(* IEC 61131-3 sources: PLC-Static-Analysis/modules/plc-rules/src/test/resources/PLCA-L008, 2 files *)

(* ---- compliant.st ---- *)
PROGRAM P_L008ok
VAR
    n : INT;
    m : INT;
    r : REAL;
    b : BOOL;
    c : BOOL;
    q : BOOL;
END_VAR
IF n > 10 THEN
    n := n - 20;
    IF n > 5 THEN
        q := TRUE;
    END_IF
END_IF
FOR m := 1 TO 10 DO
    IF n > 10 THEN
        q := TRUE;
    END_IF
    n := n + 1;
END_FOR
IF n > 10 THEN
    IF n > 50 THEN
        q := TRUE;
    END_IF
END_IF
END_PROGRAM

(* ---- noncompliant.st ---- *)
PROGRAM P_L008
VAR
    n : INT;
    m : INT;
    r : REAL;
    b : BOOL;
    c : BOOL;
    q : BOOL;
END_VAR
IF n > 10 THEN
    IF n > 5 THEN // PLCA-L008
        q := TRUE;
    END_IF
END_IF
IF m <= 0 THEN
    RETURN;
END_IF
IF m > 0 THEN // PLCA-L008
    q := TRUE;
END_IF
IF b THEN
    m := 1;
    IF b AND n > 10 THEN
        IF b THEN // PLCA-L008
            q := TRUE;
        ELSE
            q := FALSE;
        END_IF
    END_IF
END_IF
END_PROGRAM
